Staubli VAL3: setZoneFrame.pgx

public program setZoneFrame()
  local num x_nIndex
  local pointRx l_pPoint1
  local pointRx l_pPoint2
  local pointRx l_pPoint3
  local num l_nResult
begin
  link(l_pPoint1,world)
  link(l_pPoint2,world)
  link(l_pPoint3,world)
  l_pPoint1=safeTemp:zZoneItem[x_nIndex].pO
  l_pPoint2=safeTemp:zZoneItem[x_nIndex].pX
  l_pPoint3=safeTemp:zZoneItem[x_nIndex].pY
  l_nResult=setFrame(l_pPoint1,l_pPoint2,l_pPoint3,safeTemp:zZoneItem[x_nIndex].fBase)
  if l_nResult<0
    userPageAlert("坐标系生成失败："+toString("",x_nIndex))
    logMsg("坐标系生成失败："+toString("",x_nIndex))
  endIf
end
